Fanuc KAREL source: kx00026.KL

-- PROVISIONAL review KL for V1013-1; original PC SHA256 328057c7128d8ebb46db6d4a13c6aab48c5b8391d6984a13f2daea5f50651535
-- Incomplete behavior may be omitted. Consult companion uncertainty JSON. Do not deploy.
PROGRAM KX00026
%NOLOCKGROUP
VAR
  I : INTEGER
  J : INTEGER
  B : BOOLEAN
  F : FILE
  S : STRING[80]
-- UNRESOLVED_DECL P type=000102
BEGIN
  -- UNRESOLVED_PC offsets 5-12; opcodes 9D,23
  -- UNRESOLVED_PC offsets 17-21; opcodes 7F
END KX00026
